// TIA Portal V20 export
DATA_BLOCK "T4_Datos"   // DB41900
{ S7_Optimized_Access := 'TRUE' }
AUTHOR : IA
FAMILY : PRUEBA
VERSION : 0.1
// Tanda 1: datos de las pruebas
// stored: AutoNumber false
   VAR
      Tog : Bool;   // Cambia en cada ciclo (lo escribe T4_Base)
      Falso : Bool := false;   // Siempre FALSE
      Int_5 : Int := 5;   // Constante 5
      Int_3 : Int := 3;   // Constante 3
      Real_16 : Real := 16.0;   // Constante 16.0
      Real_2 : Real := 2.0;   // Constante 2.0
      Word_00F0 : Word := 16#00F0;   // Constante 16#00F0
      Word_0033 : Word := 16#0033;   // Constante 16#0033
      Mem_Runtime : LReal;
      ICoil_Q : Bool;
      SR_Mem : Bool;
      SR_Q : Bool;
      RS_Mem : Bool;
      RS_Q : Bool;
      PCont_Mem : Bool;
      NCont_Mem : Bool;
      NBox_Mem : Bool;
      PCoil_Mem : Bool;
      PCoil_Q : Bool;
      Bits_BF : Array[0..7] of Bool;
      OK_Q : Bool;
      NOTOK_Q : Bool;
      Mod_Out : Int;
      Neg_Out : Int;
      Inc_Var : Int;
      Dec_Var : Int;
      Abs_Out : Int;
      Int_m5 : Int := -5;   // Constante -5
      Min_Out : Int;
      Max_Out : Int;
      Limit_Out : Int;
      Real_2_75 : Real := 2.75;   // Constante 2.75
      Sqr_Out : Real;
      Sqrt_Out : Real;
      Ln_Out : Real;
      Exp_Out : Real;
      Sin_Out : Real;
      Cos_Out : Real;
      Tan_Out : Real;
      Frac_Out : Real;
      Real_0_5 : Real := 0.5;   // Constante 0.5
      Asin_Out : Real;
      Acos_Out : Real;
      Atan_Out : Real;
      Expt_Out : Real;
      Arr_A : Array[0..9] of Int;
      Arr_B : Array[0..9] of Int;
      Arr_C : Array[0..9] of Int;
      Arr_D : Array[0..9] of Int;
      Arr_E : Array[0..9] of Int;
      MBV_Ret : Int;
      COE_Out : UDInt;
      Arr_S1 : Array[0..9] of Int;
      Arr_S2 : Array[0..9] of Int;
      Arr_S3 : Array[0..9] of Int;
      Round_Out : DInt;
      Round_In : Real := 2.5;   // Constante 2.5
      Ceil_Out : DInt;
      Ceil_In : Real := 2.5;   // Constante 2.5
      Floor_Out : DInt;
      Floor_In : Real := 2.5;   // Constante 2.5
      Trunc_Out : DInt;
      Trunc_In : Real := 2.5;   // Constante 2.5
      ScaleX_Out : Int;
      NormX_Out : Real;
      And_Out : Word;
      Or_Out : Word;
      Xor_Out : Word;
      Inv_Out : Word;
      Deco_Out : DWord;
      Enco_Out : Int;
      Sel_Out : Int;
      Mux_Out : Int;
      Demux_0 : Int;
      Demux_1 : Int;
      Shr_Out : Word;
      Shl_Out : Word;
      Ror_Out : Word;
      Rol_Out : Word;
   END_VAR
BEGIN
END_DATA_BLOCK
